FUNCTION_BLOCK SEC_MASK_QUARTER_ACT (* Istwert (Actual CWS) mit BIT-Maske sperren: gesperrte Section 01 wird 00, Fehler und nicht installiert bleiben sichtbar *)
  (* Standard: 61499-2; Description: Copyright (c) 2026 Meisterschulen am Ostbahnhof This program and the accompanying materials are made available under the terms of the Eclipse Public License 2.0 which is available at https://www.eclipse.org/legal/epl-2.0/ SPDX-License-Identifier: EPL-2.0 *)
  (* Version 1.0, 2026-10-31, Franz Höpfinger, Meisterschulen am Ostbahnhof, initial implementation *)
  PACKAGE logiBUS::sections;
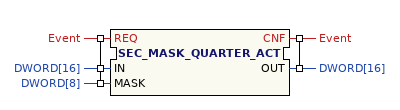
  EVENT_INPUT
    REQ WITH IN, MASK; (* Maske anwenden *)
  END_EVENT
  EVENT_OUTPUT
    CNF WITH OUT; (* Ergebnis berechnet *)
  END_EVENT
  VAR_INPUT
    IN : ARRAY [0..15] OF DWORD; (* Condensed Work State, 2 Bit je Section, Wort k = Sections 16k+1..16k+16 *)
    MASK : ARRAY [0..7] OF DWORD; (* BIT-Maske, 1 = Section frei, Wort k = Sections 32k+1..32k+32 *)
  END_VAR
  VAR_OUTPUT
    OUT : ARRAY [0..15] OF DWORD; (* Gesperrt: 01 wird 00, 00/10/11 bleiben. Frei: unveraendert *)
  END_VAR
  EC_STATES
    REQ : REQ -> CNF;
  END_STATES
  ALGORITHM REQ IN ST: (* Maske anwenden *)
VAR_TEMP
	w : UINT; // Wortindex Quarter-Array
	j : UINT; // Section im Wort
	maskWord : DWORD; // Maskenwort
	q : DWORD; // Quarter-Wert der Section
	free : BOOL; // Section laut Maske frei
	acc : DWORD; // Ergebniswort in Arbeit
END_VAR
(* Section s = 16*w + j + 1 liegt im Quarter-Array in Wort w, Bits 2j+1..2j,
   in der BIT-Maske in Wort w DIV 2, Bit 16*(w MOD 2) + j *)
FOR w := 0 TO 15 DO
	maskWord := MASK[w / 2];
	acc := DWORD#0;
	FOR j := 0 TO 15 DO
		free := (SHR(maskWord, 16 * (w MOD 2) + j) AND DWORD#1) = DWORD#1;
		q := SHR(IN[w], 2 * j) AND DWORD#2#11;
		IF free OR (q <> DWORD#2#01) THEN
			acc := acc OR SHL(q, 2 * j);
		END_IF;
	END_FOR;
	OUT[w] := acc;
END_FOR;
  END_ALGORITHM
END_FUNCTION_BLOCK
